(* IEC 61131-3 sources: PLC_ST_Simulator/examples/allgemein, 4 files *)

(* ---- Station.st ---- *)
(* Zwei Bearbeitungsstationen als Instanzen eines FB.
   Schrittkette als IF/ELSIF über nSchritt mit relativer Weiterschaltung (nSchritt := nSchritt + 10).
   Der Ablaufplan wird je Instanz erzeugt: PLC_PRG.st1.nSchritt und PLC_PRG.st2.nSchritt. *)
VAR_GLOBAL
    xStart  AT %IX0.0 : BOOL;   (* Starttaster *)
    xTeil1  AT %IX0.1 : BOOL;   (* Teil in Station 1 *)
    xB1     AT %IX0.2 : BOOL;   (* Zylinder 1 vorne *)
    xB2     AT %IX0.3 : BOOL;   (* Zylinder 1 hinten *)
    xTeil2  AT %IX0.4 : BOOL;   (* Teil in Station 2 *)
    xB3     AT %IX0.5 : BOOL;   (* Zylinder 2 vorne *)
    xB4     AT %IX0.6 : BOOL;   (* Zylinder 2 hinten *)
    xY1     AT %QX0.0 : BOOL;   (* Zylinder 1 ausfahren *)
    xY2     AT %QX0.1 : BOOL;   (* Zylinder 2 ausfahren *)
END_VAR

FUNCTION_BLOCK FB_Station
VAR_INPUT
    xStart     : BOOL;
    xTeilDa    : BOOL;
    xZylVorne  : BOOL;
    xZylHinten : BOOL;
END_VAR
VAR_OUTPUT
    xZylAus : BOOL;
    xFertig : BOOL;
END_VAR
VAR
    nSchritt : INT := 0;
    tWarte   : TON;
END_VAR

tWarte(IN := nSchritt = 30, PT := T#500MS);

IF nSchritt = 0 AND xStart AND xTeilDa THEN
    nSchritt := 10;
END_IF

IF nSchritt = 10 THEN           (* ausfahren *)
    xZylAus := TRUE;
    IF xZylVorne THEN nSchritt := nSchritt + 10; END_IF
ELSIF nSchritt = 20 THEN        (* einfahren *)
    xZylAus := FALSE;
    IF xZylHinten THEN nSchritt := 30; END_IF
ELSIF nSchritt = 30 THEN        (* warten *)
    IF tWarte.Q THEN nSchritt := 40; END_IF
ELSIF nSchritt = 40 THEN        (* fertig, Teil entnehmen *)
    xFertig := TRUE;
    IF NOT xTeilDa THEN
        xFertig := FALSE;
        nSchritt := 0;
    END_IF
END_IF
END_FUNCTION_BLOCK

PROGRAM PLC_PRG
VAR
    st1, st2 : FB_Station;
END_VAR
st1(xStart := xStart, xTeilDa := xTeil1, xZylVorne := xB1, xZylHinten := xB2, xZylAus => xY1);
st2(xStart := st1.xFertig, xTeilDa := xTeil2, xZylVorne := xB3, xZylHinten := xB4, xZylAus => xY2);
END_PROGRAM

(* ---- Ampel.st ---- *)
(* Ampel als Zustandsautomat über eine Aufzählung (CASE eZustand OF …). *)
TYPE E_Ampel : (AUS := 0, ROT, ROT_GELB, GRUEN, GELB); END_TYPE

PROGRAM PLC_PRG
VAR
  xEin AT %IX0.0 : BOOL;
  xRot AT %QX0.0 : BOOL;
  xGelb AT %QX0.1 : BOOL;
  xGruen AT %QX0.2 : BOOL;
  eZustand : E_Ampel := E_Ampel.AUS;
  tonPhase : TON;
END_VAR
tonPhase(IN := eZustand <> E_Ampel.AUS, PT := T#2S);
CASE eZustand OF
  E_Ampel.AUS:
    IF xEin THEN eZustand := E_Ampel.ROT; END_IF
  E_Ampel.ROT:
    IF tonPhase.Q THEN eZustand := E_Ampel.ROT_GELB; tonPhase(IN := FALSE); END_IF
  E_Ampel.ROT_GELB:
    IF tonPhase.Q THEN eZustand := E_Ampel.GRUEN; tonPhase(IN := FALSE); END_IF
  E_Ampel.GRUEN:
    IF tonPhase.Q THEN eZustand := E_Ampel.GELB; tonPhase(IN := FALSE); END_IF
  E_Ampel.GELB:
    IF tonPhase.Q THEN eZustand := E_Ampel.ROT; tonPhase(IN := FALSE); END_IF
END_CASE
IF NOT xEin THEN eZustand := E_Ampel.AUS; END_IF
xRot := eZustand = E_Ampel.ROT OR eZustand = E_Ampel.ROT_GELB;
xGelb := eZustand = E_Ampel.ROT_GELB OR eZustand = E_Ampel.GELB;
xGruen := eZustand = E_Ampel.GRUEN;
END_PROGRAM

(* ---- Schrittmerker.st ---- *)
(* Schrittkette aus BOOL-Schrittmerkern S0..S3: IF S1 AND xOben THEN S1 := FALSE; S2 := TRUE; END_IF *)
PROGRAM PLC_PRG
VAR
  S0 : BOOL := TRUE;
  S1, S2, S3 : BOOL;
  xStart, xOben, xUnten, xReset : BOOL;
  xMotorAuf, xMotorAb : BOOL;
END_VAR
IF S0 AND xStart THEN S0 := FALSE; S1 := TRUE; END_IF
IF S1 AND xOben THEN S1 := FALSE; S2 := TRUE; END_IF
IF S2 AND xUnten THEN S2 := FALSE; S3 := TRUE; END_IF
IF S3 AND NOT xStart THEN S3 := FALSE; S0 := TRUE; END_IF
IF xReset THEN S1 := FALSE; S2 := FALSE; S3 := FALSE; S0 := TRUE; END_IF
xMotorAuf := S1;
xMotorAb := S2;
END_PROGRAM

(* ---- Waschanlage.st ---- *)
(* Autowaschanlage (Portalwäsche)
   Ablauf: Auto einfahren → Vorwäsche → Bürsten (Hin- und Rückfahrt, Anzahl je Programm)
           → Spülen → Trocknen → Ausfahrt frei.
   Not-Halt oder Lichtschranke während der Fahrt → Störung, Quittieren → Grundstellung. *)

TYPE E_Wasch : (BEREIT, EINFAHREN, VORWAESCHE, BUERSTEN_VOR, BUERSTEN_ZURUECK, SPUELEN, TROCKNEN, AUSFAHRT, STOERUNG); END_TYPE

VAR_GLOBAL
    (* Eingänge *)
    xStartTaster   AT %IX0.0 : BOOL;   (* Münze eingeworfen / Start *)
    xProgPremium   AT %IX0.1 : BOOL;   (* Programmwahl: TRUE = Premium (3× bürsten) *)
    xAutoInPos     AT %IX0.2 : BOOL;   (* Auto steht richtig (Radsensor) *)
    xPortalVorne   AT %IX0.3 : BOOL;   (* Endschalter Portal vorne *)
    xPortalHinten  AT %IX0.4 : BOOL;   (* Endschalter Portal hinten *)
    xLichtschranke AT %IX0.5 : BOOL;   (* Person im Bereich *)
    xNotHalt       AT %IX0.6 : BOOL;   (* Öffner: TRUE = in Ordnung *)
    xQuittieren    AT %IX0.7 : BOOL;
    (* Ausgänge *)
    xAmpelRot      AT %QX0.0 : BOOL;
    xAmpelGruen    AT %QX0.1 : BOOL;
    xPortalVor     AT %QX0.2 : BOOL;
    xPortalZurueck AT %QX0.3 : BOOL;
    xBuersten      AT %QX0.4 : BOOL;
    xShampoo       AT %QX0.5 : BOOL;
    xWasser        AT %QX0.6 : BOOL;
    xGeblaese      AT %QX0.7 : BOOL;
    xStoerLampe    AT %QX1.0 : BOOL;
END_VAR

PROGRAM PLC_PRG
VAR
    eSchritt    : E_Wasch := E_Wasch.BEREIT;
    rtStart     : R_TRIG;
    tonVorwasch : TON;
    tonSpuelen  : TON;
    tonTrocknen : TON;
    tonAusfahrt : TON;
    nDurchgang  : INT;          (* gefahrene Bürstendurchgänge *)
    nSoll       : INT := 2;
    nAutosHeute : UDINT;
    tBlink      : TON;
    xBlink      : BOOL;
END_VAR

rtStart(CLK := xStartTaster);

(* Störung hat Vorrang vor allem *)
IF NOT xNotHalt OR (xLichtschranke AND (xPortalVor OR xPortalZurueck)) THEN
    eSchritt := E_Wasch.STOERUNG;
END_IF

tonVorwasch(IN := eSchritt = E_Wasch.VORWAESCHE, PT := T#4S);
tonSpuelen (IN := eSchritt = E_Wasch.SPUELEN,    PT := T#3S);
tonTrocknen(IN := eSchritt = E_Wasch.TROCKNEN,   PT := T#5S);
tonAusfahrt(IN := eSchritt = E_Wasch.AUSFAHRT AND NOT xAutoInPos, PT := T#2S);

CASE eSchritt OF
    E_Wasch.BEREIT:
        IF rtStart.Q THEN
            IF xProgPremium THEN nSoll := 3; ELSE nSoll := 2; END_IF
            nDurchgang := 0;
            eSchritt := E_Wasch.EINFAHREN;
        END_IF

    E_Wasch.EINFAHREN:
        IF xAutoInPos AND xPortalHinten AND NOT xLichtschranke THEN
            eSchritt := E_Wasch.VORWAESCHE;
        END_IF

    E_Wasch.VORWAESCHE:
        IF tonVorwasch.Q THEN eSchritt := E_Wasch.BUERSTEN_VOR; END_IF

    E_Wasch.BUERSTEN_VOR:
        IF xPortalVorne THEN eSchritt := E_Wasch.BUERSTEN_ZURUECK; END_IF

    E_Wasch.BUERSTEN_ZURUECK:
        IF xPortalHinten THEN
            nDurchgang := nDurchgang + 1;
            IF nDurchgang < nSoll THEN
                eSchritt := E_Wasch.BUERSTEN_VOR;
            ELSE
                eSchritt := E_Wasch.SPUELEN;
            END_IF
        END_IF

    E_Wasch.SPUELEN:
        IF tonSpuelen.Q THEN eSchritt := E_Wasch.TROCKNEN; END_IF

    E_Wasch.TROCKNEN:
        IF tonTrocknen.Q THEN eSchritt := E_Wasch.AUSFAHRT; END_IF

    E_Wasch.AUSFAHRT:
        IF tonAusfahrt.Q THEN
            nAutosHeute := nAutosHeute + 1;
            eSchritt := E_Wasch.BEREIT;
        END_IF

    E_Wasch.STOERUNG:
        IF xQuittieren AND xNotHalt AND NOT xLichtschranke THEN
            eSchritt := E_Wasch.BEREIT;
        END_IF
END_CASE

(* Ausgänge *)
tBlink(IN := NOT tBlink.Q, PT := T#500MS);
IF tBlink.Q THEN xBlink := NOT xBlink; END_IF

xPortalVor     := eSchritt = E_Wasch.BUERSTEN_VOR;
xPortalZurueck := eSchritt = E_Wasch.BUERSTEN_ZURUECK OR (eSchritt = E_Wasch.EINFAHREN AND NOT xPortalHinten);
xBuersten      := eSchritt = E_Wasch.BUERSTEN_VOR OR eSchritt = E_Wasch.BUERSTEN_ZURUECK;
xShampoo       := eSchritt = E_Wasch.VORWAESCHE;
xWasser        := eSchritt = E_Wasch.VORWAESCHE OR eSchritt = E_Wasch.SPUELEN;
xGeblaese      := eSchritt = E_Wasch.TROCKNEN;
xAmpelGruen    := eSchritt = E_Wasch.EINFAHREN OR eSchritt = E_Wasch.AUSFAHRT;
xAmpelRot      := NOT xAmpelGruen;
xStoerLampe    := eSchritt = E_Wasch.STOERUNG AND xBlink;
END_PROGRAM
